{attribute 'qualified_only'}
VAR_GLOBAL
	gvSwitchR1Up AT %I* : BOOL;
	gvSwitchR1Down AT %I* : BOOL;
END_VAR

(* stored: Version 1.1.0.1
   GVL gvlSwitches: Id {e769fc42-99e4-482c-9eed-c0cbd00c6def} *)
